// TwinCAT 3 PLC project PLC_LCLW
// ProgramVersion: 3.1.4026.25
// libraries:
//   Tc2_Standard, * (Beckhoff Automation GmbH)
//   Tc2_System, * (Beckhoff Automation GmbH)
// project tree:
//   GVLs/ GVL_IO.TcGVL
//   / PlcTask.TcTTO
//   POUs/ FB_Ausblasen.TcPOU, FB_Auslauf.TcPOU, FB_Auswerfer.TcPOU, FB_AuswurfBypass.TcPOU, FB_Einlauf.TcPOU, FB_Spanner.TcPOU, FB_Weiche.TcPOU, FB_ZylinderAuslauf.TcPOU, FB_ZylinderEinlauf.TcPOU, MAIN.TcPOU
// real-time tasks:
//   TASK PlcTask: cycle T#10ms, priority 20, ADS port 350
// motion (NC):
//   TASK NC-Task 1 SAF: cycle T#2ms, priority 4, ADS port 501
//   TASK NC-Task 1 SVB: cycle T#10ms, priority 8, ADS port 511
//   AXIS Axis 1 (id 1)
//     OtherSettings: AllowMotionCmdToSlave=true
//     encoder EncType=8
//       EncPara: MaxCount=#xffffffff
//     drive DrvType=9
//       DrvPara: MaxCount=#xffffffff, DriveControlDWord=#x00030100
//         Analog: VeloScale=6, TorqueSetpointScale=10, ScaleFactorActTorque=0.1
//         TimeComp: TaskDelayCycles=1
//     controller CtrType=1
//       CtrPara: PriorControlFactor=1
//         Observer: BandWidth=20
//   AXIS Axis 2 (id 2)
//     OtherSettings: AllowMotionCmdToSlave=true
//     encoder EncType=8
//       EncPara: MaxCount=#xffffffff
//     drive DrvType=9
//       DrvPara: MaxCount=#xffffffff, DriveControlDWord=#x00030100
//         Analog: VeloScale=6, TorqueSetpointScale=10, ScaleFactorActTorque=0.1
//         TimeComp: TaskDelayCycles=1
//     controller CtrType=1
//       CtrPara: PriorControlFactor=1
//         Observer: BandWidth=20
// I/O:
//   DEVICE EtherCAT_Master (disabled), AmsNetId 192.168.0.4.2.1
//     EK1100_6K1 [EK1100 EtherCAT Coupler (2A E-Bus)] (disabled)
//       EL1809_6K10 [EL1809 16Ch. Dig. Input 24V, 3ms]
//       EL2809_6K20 [EL2809 16Ch. Dig. Output 24V, 0.5A]
//     EP1018_9K1 [EP1018-0001 8 Ch. Dig. Input 24V, 10µs, M8] (disabled)
//     EP1018_9K2 [EP1018-0001 8 Ch. Dig. Input 24V, 10µs, M8] (disabled)
//     EP1018_9K3 [EP1018-0001 8 Ch. Dig. Input 24V, 10µs, M8] (disabled)
//     EP2028_10K1 [EP2028-0001 8 Ch. Dig. Output 24V, 2A, M8] (disabled)
//     EP2028_10K2 [EP2028-0001 8 Ch. Dig. Output 24V, 2A, M8] (disabled)
//     AX5206_11T1 [AX5206-0000-0210 EtherCAT Drive (SoE, 2 Ch.)] (disabled)
//     EK1100_7K1 [EK1100 EtherCAT Coupler (2A E-Bus)] (disabled)
//       EL1809_7K10 [EL1809 16Ch. Dig. Input 24V, 3ms]
//       EL2809_7K20 [EL2809 16Ch. Dig. Output 24V, 0.5A]
// variable links:
//   NC-Task 1 SAF/Axes/Axis 1 <-> EtherCAT_Master/AX5206_11T1
//     Drive/Inputs/In/nDataIn1 <-> AT 1/Following distance
//     Drive/Inputs/In/nDcOutputTime <-> InfoData/DcOutputShift
//     Drive/Inputs/In/nState1 <-> AT 1/Drive status word @bit 8
//     Drive/Inputs/In/nState2 <-> AT 1/Drive status word
//     Drive/Inputs/In/nState4 @bit 1 <-> WcState/InputToggle
//     Drive/Inputs/In/nState4 <-> WcState/WcState
//     Drive/Outputs/Out/nCtrl1 <-> MDT 1/Master control word @bit 8
//     Drive/Outputs/Out/nDataOut1 <-> MDT 1/Position command value
//     Enc/Inputs/In/nDataIn1 <-> AT 1/Position feedback 1 value
//     Enc/Inputs/In/nDcInputTime <-> InfoData/DcInputShift
//     Enc/Inputs/In/nState4 @bit 1 <-> WcState/InputToggle
//     Enc/Inputs/In/nState4 <-> WcState/WcState
//   NC-Task 1 SAF/Axes/Axis 2 <-> EtherCAT_Master/AX5206_11T1
//     Drive/Inputs/In/nDataIn1 <-> AT 2/Following distance
//     Drive/Inputs/In/nDcOutputTime <-> InfoData/DcOutputShift
//     Drive/Inputs/In/nState1 <-> AT 2/Drive status word @bit 8
//     Drive/Inputs/In/nState2 <-> AT 2/Drive status word
//     Drive/Inputs/In/nState4 @bit 1 <-> WcState/InputToggle
//     Drive/Inputs/In/nState4 <-> WcState/WcState
//     Drive/Outputs/Out/nCtrl1 <-> MDT 2/Master control word @bit 8
//     Drive/Outputs/Out/nDataOut1 <-> MDT 2/Position command value
//     Enc/Inputs/In/nDataIn1 <-> AT 2/Position feedback 1 value
//     Enc/Inputs/In/nDcInputTime <-> InfoData/DcInputShift
//     Enc/Inputs/In/nState4 @bit 1 <-> WcState/InputToggle
//     Enc/Inputs/In/nState4 <-> WcState/WcState

CONFIGURATION PLC_LCLW
    RESOURCE PLC ON TwinCAT3
        TASK PlcTask(INTERVAL := T#10ms, PRIORITY := 20);
        PROGRAM MAIN WITH PlcTask : MAIN;
    END_RESOURCE
END_CONFIGURATION

// ---- GVLs/GVL_IO.TcGVL
{attribute 'qualified_only'}
VAR_GLOBAL
	 xNotHalt_Betaetigt : BOOL;           // E0.1 - Not-Halt betätigt 
     xLaserEnable : BOOL;                 // A0.1 - LaserEnable
	 xLichtschranke_Einlauf : BOOL;       // E1052.0 - Lichtschranke Einlauf
     xServo_Einlauf_Eingerastet : BOOL;   // E1052.1 - Servo Einlauf eingerastet
     xServo_Einlauf_AS : BOOL;            // E1052.2 - Servo Einlauf AS
     xServo_Einlauf_GS : BOOL;            // E1052.3 - Servo Einlauf GS
	 xEinlaufBereit : BOOL;               // Part ready at infeed (calculated, not a direct sensor)
	 xZylinderSpannerAS : BOOL;           // E1050.2 - Zylinder Spanner AS
     xZylinderSpannerGS : BOOL;           // E1050.3 - Zylinder Spanner GS
     xVentilSpannerAS : BOOL;             // A1050.2 - Ventil Spanner AS
     xVentilSpannerGS : BOOL;             // A1050.3 - Ventil Spanner GS
	 xZylinderEinlaufAS : BOOL;           // E1051.0 - Zylinder Einlauf AS
     xZylinderEinlaufGS : BOOL;           // E1051.1 - Zylinder Einlauf GS
     xVentilEinlaufAS : BOOL;             // A1051.0 - Ventil Einlauf AS
     xVentilEinlaufGS : BOOL;             // A1051.1 - Ventil Einlauf GS
     xZylinderEinlaufBereit : BOOL;       // Calculated: cylinder confirmed in position
	 xSpannerBereit : BOOL;               // Calculated: clamp confirmed closed (from E1050.2 feedback)
     xPartOK : BOOL;                      // PLACEHOLDER: simulated quality decision, normally from an external vision/quality system not present in this Eplan/pneumatic scope — forced manually for testing
     xZylinderWeicheAS : BOOL;   // E1050.4 - Zylinder Weiche AS
     xZylinderWeicheGS : BOOL;   // E1050.5 - Zylinder Weiche GS
     xVentilWeicheAS : BOOL;     // A1050.4 - Ventil Weiche AS
     xVentilWeicheGS : BOOL;     // A1050.5 - Ventil Weiche GS
     xWeicheRejectBereit : BOOL; // Calculated: diverter confirmed in reject position
     xWeicheAcceptBereit : BOOL; // Calculated: diverter confirmed in accept/straight position
	 xZylinderAuswerferAS : BOOL;   // E1050.0 - Zylinder Auswerfer AS
     xZylinderAuswerferGS : BOOL;   // E1050.1 - Zylinder Auswerfer GS
     xVentilAuswerferAS : BOOL;     // A1050.0 - Ventil Auswerfer AS
     xVentilAuswerferGS : BOOL;     // A1050.1 - Ventil Auswerfer GS
     xVentilAusblasenAS : BOOL;     // A1051.4 - Ventil Ausblasen AS
     xVentilAusblasenGS : BOOL;     // A1051.5 - Ventil Ausblasen GS
     xAuswerferBereit : BOOL;       // Calculated: ejector confirmed extended
	 xZylinderAuslaufAS : BOOL;     // E1051.2 - Zylinder Auslauf AS
     xZylinderAuslaufGS : BOOL;     // E1051.3 - Zylinder Auslauf GS
     xVentilAuslaufAS : BOOL;       // A1051.2 - Ventil Auslauf AS
     xVentilAuslaufGS : BOOL;       // A1051.3 - Ventil Auslauf GS
     xZylinderAuslaufBereit : BOOL; // Calculated: outfeed cylinder confirmed in position

     xLichtschranke_Auslauf : BOOL;       // E1052.4 - Lichtschranke Auslauf
     xServo_Auslauf_Eingerastet : BOOL;   // E1052.5 - Servo Auslauf eingerastet
     xServo_Auslauf_AS : BOOL;            // E1052.6 - Servo Auslauf AS
	 xServo_Auslauf_GS : BOOL;            // E1052.7 - Servo Auslauf GS
	 xAuslaufBereit : BOOL;               // Calculated: part confirmed exited

	 xVentilAuswurfBypassAS : BOOL;   // A1051.6 - Ventil Auswurf Bypass AS
	 xVentilAuswurfBypassGS : BOOL;   // A1051.7 - Ventil Auswurf Bypass GS
	 xBypassTrigger : BOOL;   // PLACEHOLDER: no defining condition exists in either drawing, forced manually for testing
END_VAR

// ---- POUs/MAIN.TcPOU
PROGRAM MAIN
VAR
    fbEinlauf : FB_Einlauf;
	fbZylinderEinlauf : FB_ZylinderEinlauf;
    fbSpanner : FB_Spanner;
	fbWeiche : FB_Weiche;
	fbAuswerfer : FB_Auswerfer;
    fbAusblasen : FB_Ausblasen;
	fbZylinderAuslauf : FB_ZylinderAuslauf;
    fbAuslauf : FB_Auslauf;
    fbAuswurfBypass : FB_AuswurfBypass;
END_VAR

GVL_IO.xLaserEnable := NOT GVL_IO.xNotHalt_Betaetigt;
fbEinlauf();
fbZylinderEinlauf();
fbSpanner();
fbWeiche();
fbAuswerfer();
fbAusblasen();
fbZylinderAuslauf();
fbAuslauf();
fbAuswurfBypass();

END_PROGRAM

// ---- POUs/FB_Einlauf.TcPOU
FUNCTION_BLOCK FB_Einlauf
VAR_INPUT
END_VAR
VAR_OUTPUT
END_VAR
VAR
END_VAR

IF GVL_IO.xLichtschranke_Einlauf AND GVL_IO.xServo_Einlauf_GS THEN
    GVL_IO.xEinlaufBereit := TRUE;
ELSIF NOT GVL_IO.xLichtschranke_Einlauf THEN
    GVL_IO.xEinlaufBereit := FALSE;
END_IF

END_FUNCTION_BLOCK

// ---- POUs/FB_ZylinderEinlauf.TcPOU
FUNCTION_BLOCK FB_ZylinderEinlauf
VAR_INPUT
END_VAR
VAR_OUTPUT
END_VAR
VAR
END_VAR

GVL_IO.xVentilEinlaufAS := GVL_IO.xEinlaufBereit;
GVL_IO.xVentilEinlaufGS := NOT GVL_IO.xEinlaufBereit;
GVL_IO.xZylinderEinlaufBereit := GVL_IO.xZylinderEinlaufAS;

END_FUNCTION_BLOCK

// ---- POUs/FB_Spanner.TcPOU
FUNCTION_BLOCK FB_Spanner
VAR_INPUT
END_VAR
VAR_OUTPUT
END_VAR
VAR
END_VAR

GVL_IO.xVentilSpannerAS := GVL_IO.xZylinderEinlaufBereit;
GVL_IO.xVentilSpannerGS := NOT GVL_IO.xZylinderEinlaufBereit;
GVL_IO.xSpannerBereit := GVL_IO.xZylinderSpannerAS;

END_FUNCTION_BLOCK

// ---- POUs/FB_Weiche.TcPOU
FUNCTION_BLOCK FB_Weiche
VAR_INPUT
END_VAR
VAR_OUTPUT
END_VAR
VAR
END_VAR

GVL_IO.xVentilWeicheAS := GVL_IO.xSpannerBereit AND NOT GVL_IO.xPartOK;
GVL_IO.xVentilWeicheGS := GVL_IO.xSpannerBereit AND GVL_IO.xPartOK;

GVL_IO.xWeicheRejectBereit := GVL_IO.xZylinderWeicheAS;
GVL_IO.xWeicheAcceptBereit := GVL_IO.xZylinderWeicheGS;

END_FUNCTION_BLOCK

// ---- POUs/FB_Auswerfer.TcPOU
FUNCTION_BLOCK FB_Auswerfer
VAR_INPUT
END_VAR
VAR_OUTPUT
END_VAR
VAR
END_VAR

GVL_IO.xVentilAuswerferAS := GVL_IO.xWeicheRejectBereit;
GVL_IO.xVentilAuswerferGS := NOT GVL_IO.xWeicheRejectBereit;

GVL_IO.xAuswerferBereit := GVL_IO.xZylinderAuswerferAS;

END_FUNCTION_BLOCK

// ---- POUs/FB_Ausblasen.TcPOU
FUNCTION_BLOCK FB_Ausblasen
VAR_INPUT
END_VAR
VAR_OUTPUT
END_VAR
VAR
tonBlow : TON;
END_VAR

tonBlow(IN := GVL_IO.xAuswerferBereit, PT := T#1S);

GVL_IO.xVentilAusblasenAS := GVL_IO.xAuswerferBereit AND NOT tonBlow.Q;
GVL_IO.xVentilAusblasenGS := NOT GVL_IO.xVentilAusblasenAS;

END_FUNCTION_BLOCK

// ---- POUs/FB_ZylinderAuslauf.TcPOU
FUNCTION_BLOCK FB_ZylinderAuslauf
VAR_INPUT
END_VAR
VAR_OUTPUT
END_VAR
VAR
END_VAR

GVL_IO.xVentilAuslaufAS := GVL_IO.xWeicheAcceptBereit;
GVL_IO.xVentilAuslaufGS := NOT GVL_IO.xWeicheAcceptBereit;

GVL_IO.xZylinderAuslaufBereit := GVL_IO.xZylinderAuslaufAS;

END_FUNCTION_BLOCK

// ---- POUs/FB_Auslauf.TcPOU
FUNCTION_BLOCK FB_Auslauf
VAR_INPUT
END_VAR
VAR_OUTPUT
END_VAR
VAR
END_VAR

IF GVL_IO.xLichtschranke_Auslauf AND GVL_IO.xServo_Auslauf_GS THEN
    GVL_IO.xAuslaufBereit := TRUE;
ELSIF NOT GVL_IO.xLichtschranke_Auslauf THEN
    GVL_IO.xAuslaufBereit := FALSE;
END_IF

END_FUNCTION_BLOCK

// ---- POUs/FB_AuswurfBypass.TcPOU
FUNCTION_BLOCK FB_AuswurfBypass
VAR_INPUT
END_VAR
VAR_OUTPUT
END_VAR
VAR
	tonBypass : TON;
END_VAR

tonBypass(IN := GVL_IO.xBypassTrigger, PT := T#1S);

GVL_IO.xVentilAuswurfBypassAS := GVL_IO.xBypassTrigger AND NOT tonBypass.Q;
GVL_IO.xVentilAuswurfBypassGS := NOT GVL_IO.xVentilAuswurfBypassAS;

END_FUNCTION_BLOCK
